// TwinCAT 3 PLC project FillPlc
// ProgramVersion: 3.1.4026.12
// project tree:
//   DUTs/ E_FillState.TcDUT, ST_Recipe.TcDUT
//   GVLs/ GVL_IO.TcGVL, GVL_Alarms.TcGVL
//   POUs/ FB_Valve.TcPOU, FB_Device.TcPOU, FB_Pump.TcPOU, F_Scale.TcPOU, MAIN.TcPOU
//   / PlcTask.TcTTO

CONFIGURATION FillPlc
    RESOURCE PLC ON TwinCAT3
        TASK PlcTask(INTERVAL := T#10ms, PRIORITY := 20);
        PROGRAM MAIN WITH PlcTask : MAIN;
    END_RESOURCE
END_CONFIGURATION

// ---- DUTs/E_FillState.TcDUT
// Steps of the fill sequence
{attribute 'qualified_only'}
{attribute 'strict'}
TYPE E_FillState :
(
	Idle := 0,        // waiting for Start
	Filling := 10,    // inlet valve open
	Settling := 20,
	Draining := 30,
	Fault := 99
) INT;
END_TYPE

// ---- DUTs/ST_Recipe.TcDUT
TYPE ST_Recipe :
STRUCT
	fLevelSetpoint : REAL := 80.0;   // fill level to reach in %
	tSettle : TIME := T#5S;          // how long the product settles
	(* recipe number from MES *)
	nRecipeNo : DINT;
	sName : STRING(40);
END_STRUCT
END_TYPE

// ---- GVLs/GVL_IO.TcGVL
// Field inputs and outputs, linked to the EtherCAT terminals
{attribute 'qualified_only'}
VAR_GLOBAL
	bStartButton AT %I* : BOOL;      // Start push button S1
	bStopButton AT %I* : BOOL;       // Stop push button S2 (NC)
	bInletOpen AT %I* : BOOL;        // XV1 open limit switch
	nLevelRaw AT %I* : INT;          // LT1 level, raw 0..32767
	bInletValve AT %Q* : BOOL;       // XV1 inlet valve solenoid
	bPumpRun AT %Q* : BOOL;          // P1 drain pump contactor
END_VAR
VAR_GLOBAL CONSTANT
	cMaxLevel : REAL := 95.0;
END_VAR

// ---- GVLs/GVL_Alarms.TcGVL
VAR_GLOBAL
	aAlarm : ARRAY[1..4] OF BOOL;   // 1 XV1 not open, 2 level high-high, 3 pump fault, 4 fill timeout
	bAnyFault : BOOL;
END_VAR

// ---- POUs/MAIN.TcPOU
PROGRAM MAIN
VAR
	eState : E_FillState;          // fill sequence step
	fLevel : REAL;                 // tank level LT1 in %
	stRecipe : ST_Recipe;
	fbInlet : FB_Valve;            // XV1 inlet valve
	fbDrain : FB_Pump;             // P1 drain pump
	tonStep : TON;                 // time in step
	(* "Stop" pressed: wait for Start *)
	bPaused : BOOL;
END_VAR

// level from the analog input
fLevel := F_Scale(nRaw := GVL_IO.nLevelRaw, fMax := 100.0);

IF NOT GVL_IO.bStopButton THEN
	bPaused := TRUE;
ELSIF GVL_IO.bStartButton THEN
	bPaused := FALSE;
END_IF

CASE eState OF
	E_FillState.Idle:
		IF GVL_IO.bStartButton AND NOT GVL_Alarms.bAnyFault THEN
			eState := E_FillState.Filling;
		END_IF
	E_FillState.Filling:
		IF fLevel >= stRecipe.fLevelSetpoint THEN
			eState := E_FillState.Settling;
		END_IF
	E_FillState.Settling:
		IF tonStep.Q THEN
			eState := E_FillState.Draining;
		END_IF
	E_FillState.Draining:
		IF fLevel < 2.0 THEN
			eState := E_FillState.Idle;
		END_IF
END_CASE
tonStep(IN := eState = E_FillState.Settling, PT := stRecipe.tSettle);

fbInlet(bOpenReq := eState = E_FillState.Filling AND NOT bPaused,
        bPermit := fLevel < GVL_IO.cMaxLevel,
        bOpenFb := GVL_IO.bInletOpen);
GVL_IO.bInletValve := fbInlet.bOpenCmd;

fbDrain(bRunReq := eState = E_FillState.Draining);
GVL_IO.bPumpRun := fbDrain.bRunCmd;

GVL_Alarms.aAlarm[1] := fbInlet.bFaultNotOpen;
GVL_Alarms.bAnyFault := GVL_Alarms.aAlarm[1] OR GVL_Alarms.aAlarm[2] OR GVL_Alarms.aAlarm[3];

END_PROGRAM

// ---- POUs/FB_Valve.TcPOU
// On/off valve with open feedback and travel monitoring
FUNCTION_BLOCK FB_Valve
VAR_INPUT
	bOpenReq : BOOL;          // program wants the valve open
	bPermit : BOOL;           // interlocks OK
	bOpenFb : BOOL;           // open limit switch
	tTravel : TIME := T#10S;  // max travel time
END_VAR
VAR_OUTPUT
	bOpenCmd : BOOL;          // solenoid output
	bFaultNotOpen : BOOL;     // did not open within tTravel
END_VAR
VAR
	tonTravel : TON;
END_VAR

bOpenCmd := bOpenReq AND bPermit;
tonTravel(IN := bOpenCmd AND NOT bOpenFb, PT := tTravel);
IF tonTravel.Q THEN
	bFaultNotOpen := TRUE;
END_IF

METHOD Reset : BOOL
bFaultNotOpen := FALSE;
END_METHOD

END_FUNCTION_BLOCK

// ---- POUs/FB_Pump.TcPOU
FUNCTION_BLOCK FB_Pump EXTENDS FB_Device
VAR_INPUT
	bRunReq : BOOL;   // program wants the pump running
END_VAR
VAR_OUTPUT
	bRunCmd : BOOL;   // contactor output
END_VAR

bRunCmd := bRunReq AND NOT bFault;

END_FUNCTION_BLOCK

// ---- POUs/FB_Device.TcPOU
FUNCTION_BLOCK ABSTRACT FB_Device
VAR_OUTPUT
	bFault : BOOL;   // device fault
END_VAR

END_FUNCTION_BLOCK

// ---- POUs/F_Scale.TcPOU
// Raw analog value to engineering units
FUNCTION F_Scale : REAL
VAR_INPUT
	nRaw : INT;
	fMax : REAL;
END_VAR
VAR
	fTmp : REAL;
END_VAR

fTmp := INT_TO_REAL(nRaw) / 32767.0;
F_Scale := fTmp * fMax;

END_FUNCTION
